// TIA Portal V21 export
// export: Created 2026-11-11T00:47:17.260442Z, ExportSetting WithDefaults, DisplayName Totally Integrated Automation Portal, DisplayVersion V21 Update 3, DisplayName STEP 7 Professional, DisplayVersion V21 Update 3, DisplayName STEP 7 Safety, DisplayVersion V21, DisplayName Tech WebApplication, DisplayVersion V21, DisplayName WinCC Basic/Comfort/Advanced, DisplayVersion V21 Update 3, DisplayName WinCC Unified, DisplayVersion V21 Update 3
FUNCTION_BLOCK "FB_Fbd_ex045"   // FB88, FBD
{ S7_Optimized_Access := 'TRUE' }
VERSION : 0.1
// stored: AutoNumber true, IsIECCheckEnabled false, IsRetainMemResEnabled false, MemoryReserve 100, SetENOAutomatically false, UDAEnableTagReadback false
   VAR_INPUT
      v_req : Bool;
      v_id : HW_IO;
      v_index : DInt;
      v_mlen : UInt;
   END_VAR
   VAR_OUTPUT
      v_valid : Bool;
      v_busy : Bool;
      v_error : Bool;
      v_status : DWord;
      v_len : UInt;
   END_VAR
   VAR_IN_OUT
      v_record : Array[0..99] of Byte;
   END_VAR
   VAR
      inst { S7_SetPoint := 'True'} : RDREC;
   END_VAR
BEGIN

REGION Network 1: RDREC - Read data record
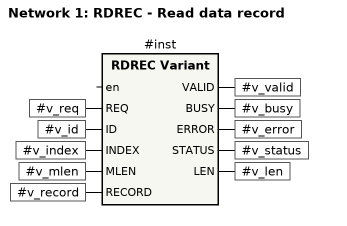
   #inst(REQ := #v_req,   // RDREC
         ID := #v_id,
         INDEX := #v_index,
         MLEN := #v_mlen,
         RECORD := #v_record,
         VALID => #v_valid,
         BUSY => #v_busy,
         ERROR => #v_error,
         STATUS => #v_status,
         LEN => #v_len);
END_REGION
END_FUNCTION_BLOCK
